ABB RAPID module: test.modx

MODULE A1_457_L
    ! ----------------------------------------------------------------------
    ! Robot ABB serial n. IRB  6720-101047
    ! ----------------------------------------------------------------------
    ! Final customer :  Martin Rea
    ! ----------------------------------------------------------------------
    ! Cell made by :    TREBI - Cellatica (BS) - Italy
    ! ----------------------------------------------------------------------
    ! Job order n. :    21301
    ! ----------------------------------------------------------------------
    ! Programmer :      Turati Simone
    ! ----------------------------------------------------------------------
    ! Date Rev.0:       07/10/2026
    ! Date Rev.1:
    ! Date Rev.2:
    ! Date Rev.3:
    ! Date Rev.4:
    ! ----------------------------------------------------------------------
    ! +-+-+-+-+-+-+-+-+-+-+-+-+-+-+-+-+-+-+-+-+-+-+-+-+-+-+-+-+-+-+-+-+-+-+-
    ! +-+-+-+-+-+-+-+-+-+-+-+-+-+-+-+-+-+-+-+-+-+-+-+-+-+-+-+-+-+-+-+-+-+-+-
    ! +-+-+-+-+-+-+-+-+-+-+-+-+-+-+-+-+-+-+-+-+-+-+-+-+-+-+-+-+-+-+-+-+-+-+-
    !EXCHANGE DATA (Variables with "M")
    ! **********************************************************************
    ! NUM DATA
    ! **********************************************************************
    PERS num nMProg:=1;
    ! **********************************************************************
    ! STRING DATA
    ! **********************************************************************
    !Stringhe nome programma
    PERS String sMProgramName:="PART_0001";
    PERS String sMPartName:="PEZZO 1";
    ! +-+-+-+-+-+-+-+-+-+-+-+-+-+-+-+-+-+-+-+-+-+-+-+-+-+-+-+-+-+-+-+-+-+-+-
    ! +-+-+-+-+-+-+-+-+-+-+-+-+-+-+-+-+-+-+-+-+-+-+-+-+-+-+-+-+-+-+-+-+-+-+-
    ! +-+-+-+-+-+-+-+-+-+-+-+-+-+-+-+-+-+-+-+-+-+-+-+-+-+-+-+-+-+-+-+-+-+-+-
    ! **********************************************************************
    ! NUM DATA
    ! **********************************************************************
    PERS dnum nLPartCounter:=19;
    ! **********************************************************************
    ! TOOL DATA
    ! **********************************************************************
    PERS tooldata tGripp_1:=[TRUE,[[0,250,335],[1,0,0,0]],[61.3,[54,3.3,163.7],[1,0,0,0],4.49,1.158,5.024]];
    ! **********************************************************************
    ! LOAD DATA
    ! **********************************************************************
    PERS loaddata LoadPart_L:=[4.5,[16.9,32.5,271],[1,0,0,0],0.7,0.6,0.2];
    ! **********************************************************************
    ! SPEED DATA
    ! **********************************************************************
    LOCAL PERS speeddata vPicking:=[60,500,0,0];
    LOCAL PERS speeddata vUnload:=[150,500,0,0];
    LOCAL PERS speeddata vGrind1:=[200,100,0,0];
    LOCAL PERS speeddata vGrind2:=[170,80,0,0];
    ! **********************************************************************
    ! ROBTARGET DATA
    ! **********************************************************************
    ! LOAD BELT
    PERS robtarget pLAppPick:=[[800,1370,1180],[0,0.642788,-0.766044,0],[0,0,-1,0],[9E+09,9E+09,9E+09,9E+09,9E+09,9E+09]];
    PERS robtarget pLPick:=[[3.81937,161.237,727.32],[0.138322,-0.983291,0.0782176,0.0888119],[0,-1,0,0],[9E+09,9E+09,9E+09,9E+09,9E+09,9E+09]];
    PERS robtarget pLPick_0:=[[97.94,1368.66,727.32],[0.160804,-0.644231,0.746958,-0.0340974],[0,-1,0,0],[9E+09,9E+09,9E+09,9E+09,9E+09,9E+09]];
    PERS robtarget pLCHK_Part:=[[-4.50,1321.99,1326.48],[0.156146,0.631329,-0.73609,-0.187653],[0,0,-1,0],[9E+09,9E+09,9E+09,9E+09,9E+09,9E+09]];
    ! RECENTRE
    PERS robtarget pLAppRec_:=[[890,-790,1800],[0,0,0.70711,-0.70711],[-1,-2,0,0],[9E+09,9E+09,9E+09,9E+09,9E+09,9E+09]];
    PERS robtarget pLRecentre_:=[[860,-495,2540],[0,0,0,1],[-1,-2,0,0],[9E+09,9E+09,9E+09,9E+09,9E+09,9E+09]];
    ! DATAMATRIX
    PERS robtarget pLAppDataMatrix_:=[[640.77,1371.32,1306.69],[0.400689,0.173653,-0.899217,0.0265008],[0,0,0,0],[9E+09,9E+09,9E+09,9E+09,9E+09,9E+09]];
    PERS robtarget pLDataMatrix:=[[-260,1005,1305],[0.407608,0.15668,-0.89732,0.0642135],[0,0,0,0],[9E+09,9E+09,9E+09,9E+09,9E+09,9E+09]];
    ! **********************************************************************
    ! CHANGE POINT
    PERS robtarget pLAppChange_1:=[[1370,1085,1560],[0,0,-0.707107,-0.707107],[0,1,-1,0],[9E+09,9E+09,9E+09,9E+09,9E+09,9E+09]];
    PERS robtarget pLAppChange_2:=[[1370,1085,1560],[0,0,-0.707107,-0.707107],[0,1,-1,0],[9E+09,9E+09,9E+09,9E+09,9E+09,9E+09]];
    PERS robtarget pLAppChange_3:=[[1370,1085,1560],[0,0,-0.707107,-0.707107],[0,1,-1,0],[9E+09,9E+09,9E+09,9E+09,9E+09,9E+09]];
    PERS robtarget pLAppChange_4:=[[1370,1085,1560],[0,0,-0.707107,-0.707107],[0,1,-1,0],[9E+09,9E+09,9E+09,9E+09,9E+09,9E+09]];
    PERS robtarget pLAppChange_5:=[[1370,1085,1560],[0,0,-0.707107,-0.707107],[0,1,-1,0],[9E+09,9E+09,9E+09,9E+09,9E+09,9E+09]];
    PERS robtarget pLAppChange_6:=[[1370,1085,1560],[0,0,-0.707107,-0.707107],[0,1,-1,0],[9E+09,9E+09,9E+09,9E+09,9E+09,9E+09]];
    PERS robtarget pLAppChange_7:=[[1370,1085,1560],[0,0,-0.707107,-0.707107],[0,1,-1,0],[9E+09,9E+09,9E+09,9E+09,9E+09,9E+09]];
    PERS robtarget pLAppChange_8:=[[1370,1085,1560],[0,0,-0.707107,-0.707107],[0,1,-1,0],[9E+09,9E+09,9E+09,9E+09,9E+09,9E+09]];
    PERS robtarget pLAppChange_9:=[[1370,1085,1560],[0,0,-0.707107,-0.707107],[0,1,-1,0],[9E+09,9E+09,9E+09,9E+09,9E+09,9E+09]];
    PERS robtarget pLAppChange_10:=[[1370,1085,1560],[0,0,-0.707107,-0.707107],[0,1,-1,0],[9E+09,9E+09,9E+09,9E+09,9E+09,9E+09]];
    PERS robtarget pLChange:=[[1590,1800,1695],[0,0,0.707107,0.707107],[0,1,-1,0],[9E+09,9E+09,9E+09,9E+09,9E+09,9E+09]];
    ! **********************************************************************
    !Safe Homing
    PERS robtarget pLSafeHoming_OP010_:=[[0,0,0],[0,0,0,0],[0,0,0,0],[9E+09,9E+09,9E+09,9E+09,9E+09,9E+09]];
    PERS robtarget pLSafeHoming_OP020_:=[[0,0,0],[0,0,0,0],[0,0,0,0],[9E+09,9E+09,9E+09,9E+09,9E+09,9E+09]];
    PERS robtarget pLSafeHoming_OP030_:=[[0,0,0],[0,0,0,0],[0,0,0,0],[9E+09,9E+09,9E+09,9E+09,9E+09,9E+09]];
    PERS robtarget pLSafeHoming_OP040_:=[[0,0,0],[0,0,0,0],[0,0,0,0],[9E+09,9E+09,9E+09,9E+09,9E+09,9E+09]];
    PERS robtarget pLSafeHoming_OP050_:=[[0,0,0],[0,0,0,0],[0,0,0,0],[9E+09,9E+09,9E+09,9E+09,9E+09,9E+09]];
    PERS robtarget pLSafeHoming_OP060_:=[[0,0,0],[0,0,0,0],[0,0,0,0],[9E+09,9E+09,9E+09,9E+09,9E+09,9E+09]];
    PERS robtarget pLSafeHoming_OP070_:=[[0,0,0],[0,0,0,0],[0,0,0,0],[9E+09,9E+09,9E+09,9E+09,9E+09,9E+09]];
    PERS robtarget pLSafeHoming_OP080_:=[[0,0,0],[0,0,0,0],[0,0,0,0],[9E+09,9E+09,9E+09,9E+09,9E+09,9E+09]];
    PERS robtarget pLSafeHoming_OP090_:=[[0,0,0],[0,0,0,0],[0,0,0,0],[9E+09,9E+09,9E+09,9E+09,9E+09,9E+09]];
    PERS robtarget pLSafeHoming_OP100_:=[[0,0,0],[0,0,0,0],[0,0,0,0],[9E+09,9E+09,9E+09,9E+09,9E+09,9E+09]];
    PERS robtarget pLSafeHoming_OP110_:=[[0,0,0],[0,0,0,0],[0,0,0,0],[9E+09,9E+09,9E+09,9E+09,9E+09,9E+09]];
    PERS robtarget pLSafeHoming_OP120_:=[[0,0,0],[0,0,0,0],[0,0,0,0],[9E+09,9E+09,9E+09,9E+09,9E+09,9E+09]];
    PERS robtarget pLSafeHoming_OP130_:=[[0,0,0],[0,0,0,0],[0,0,0,0],[9E+09,9E+09,9E+09,9E+09,9E+09,9E+09]];
    PERS robtarget pLSafeHoming_OP140_:=[[0,0,0],[0,0,0,0],[0,0,0,0],[9E+09,9E+09,9E+09,9E+09,9E+09,9E+09]];
    PERS robtarget pLSafeHoming_OP150_:=[[0,0,0],[0,0,0,0],[0,0,0,0],[9E+09,9E+09,9E+09,9E+09,9E+09,9E+09]];
    PERS robtarget pLSafeHoming_OP160_:=[[0,0,0],[0,0,0,0],[0,0,0,0],[9E+09,9E+09,9E+09,9E+09,9E+09,9E+09]];
    PERS robtarget pLSafeHoming_OP170_:=[[0,0,0],[0,0,0,0],[0,0,0,0],[9E+09,9E+09,9E+09,9E+09,9E+09,9E+09]];
    PERS robtarget pLSafeHoming_OP180_:=[[0,0,0],[0,0,0,0],[0,0,0,0],[9E+09,9E+09,9E+09,9E+09,9E+09,9E+09]];
    PERS robtarget pLSafeHoming_OP190_:=[[0,0,0],[0,0,0,0],[0,0,0,0],[9E+09,9E+09,9E+09,9E+09,9E+09,9E+09]];
    PERS robtarget pLSafeHoming_OP200_:=[[0,0,0],[0,0,0,0],[0,0,0,0],[9E+09,9E+09,9E+09,9E+09,9E+09,9E+09]];
    ! **********************************************************************
    ! GRINDER 1
    ! **********************************************************************
    !OPXXX
    PERS robtarget pLU1_OPXXX_000:=[[0,0,0],[0,0,0,0],[0,0,0,0],[9E+09,9E+09,9E+09,9E+09,9E+09,9E+09]];
    PERS robtarget pLU1_OPXXX_010:=[[0,0,0],[0,0,0,0],[0,0,0,0],[9E+09,9E+09,9E+09,9E+09,9E+09,9E+09]];
    PERS robtarget pLU1_OPXXX_020:=[[0,0,0],[0,0,0,0],[0,0,0,0],[9E+09,9E+09,9E+09,9E+09,9E+09,9E+09]];
    PERS robtarget pLU1_OPXXX_030:=[[0,0,0],[0,0,0,0],[0,0,0,0],[9E+09,9E+09,9E+09,9E+09,9E+09,9E+09]];
    ! **********************************************************************
    ! GRINDER 2
    ! **********************************************************************
    !OP10
    PERS robtarget pLU2_OP10_000 := [[-512.78,-45.67,-339.98],[0.753965,0.177077,0.558855,-0.296414],[-1,1,2,0],[9E+09,9E+09,9E+09,9E+09,9E+09,9E+09]];
    PERS robtarget pLU2_OP10_010 := [[83.19,99.41,-382.48],[0.834702,0.222849,0.429026,-0.263719],[-1,2,2,0],[9E+09,9E+09,9E+09,9E+09,9E+09,9E+09]];
    PERS robtarget pLU2_OP10_020 := [[166.56,99.41,-332.86],[0.834697,0.222853,0.429032,-0.26372],[-1,2,2,0],[9E+09,9E+09,9E+09,9E+09,9E+09,9E+09]];
    PERS robtarget pLU2_OP10_030 := [[166.56,99.41,-309.01],[0.834699,0.222852,0.42903,-0.26372],[-1,2,2,0],[9E+09,9E+09,9E+09,9E+09,9E+09,9E+09]];
    PERS robtarget pLU2_OP10_040 := [[147.76,53.29,-309.01],[0.834699,0.222851,0.429031,-0.26372],[-1,2,2,0],[9E+09,9E+09,9E+09,9E+09,9E+09,9E+09]];
    PERS robtarget pLU2_OP10_050 := [[99.74,9.11,-312.84],[0.834697,0.222851,0.429033,-0.26372],[-1,2,2,0],[9E+09,9E+09,9E+09,9E+09,9E+09,9E+09]];
    PERS robtarget pLU2_OP10_060 := [[89.03,-30.27,-311.48],[0.834674,0.222871,0.429035,-0.263775],[-1,2,2,0],[9E+09,9E+09,9E+09,9E+09,9E+09,9E+09]];
    PERS robtarget pLU2_OP10_070 := [[89.03,-66.46,-311.47],[0.834674,0.222871,0.429033,-0.263777],[-1,2,2,0],[9E+09,9E+09,9E+09,9E+09,9E+09,9E+09]];
    PERS robtarget pLU2_OP10_080 := [[78.00,-94.61,-311.47],[0.86058,0.168979,0.452974,-0.160198],[-1,1,2,0],[9E+09,9E+09,9E+09,9E+09,9E+09,9E+09]];
    PERS robtarget pLU2_OP10_090 := [[48.43,-125.73,-310.69],[0.86058,0.168979,0.452973,-0.160199],[-1,1,2,0],[9E+09,9E+09,9E+09,9E+09,9E+09,9E+09]];
    PERS robtarget pLU2_OP10_100 := [[48.68,-150.17,-329.57],[0.86058,0.168977,0.452973,-0.160199],[-1,1,2,0],[9E+09,9E+09,9E+09,9E+09,9E+09,9E+09]];
    PERS robtarget pLU2_OP10_110 := [[-99.73,-229.10,-399.55],[0.860581,0.168977,0.452973,-0.160199],[-1,1,2,0],[9E+09,9E+09,9E+09,9E+09,9E+09,9E+09]];
    !OP20
    PERS robtarget pLU2_OP20_000 := [[-385.23,300.06,-127.42],[0.574393,0.0777966,0.781268,-0.231604],[-1,1,2,0],[9E+09,9E+09,9E+09,9E+09,9E+09,9E+09]];
    PERS robtarget pLU2_OP20_010 := [[9.44,300.13,-103.22],[0.574395,0.0777988,0.781267,-0.231602],[-1,1,2,0],[9E+09,9E+09,9E+09,9E+09,9E+09,9E+09]];
    PERS robtarget pLU2_OP20_020 := [[101.46,300.12,-56.96],[0.574396,0.0778002,0.781266,-0.231603],[-1,1,2,0],[9E+09,9E+09,9E+09,9E+09,9E+09,9E+09]];
    PERS robtarget pLU2_OP20_030 := [[101.45,300.13,-43.36],[0.574393,0.0778009,0.781269,-0.231601],[-1,1,2,0],[9E+09,9E+09,9E+09,9E+09,9E+09,9E+09]];
    PERS robtarget pLU2_OP20_040 := [[101.45,261.09,-43.36],[0.574393,0.0778004,0.781269,-0.231601],[-1,1,2,0],[9E+09,9E+09,9E+09,9E+09,9E+09,9E+09]];
    PERS robtarget pLU2_OP20_050 := [[83.98,199.96,-132.65],[0.51864,-0.0749808,0.781563,-0.338452],[-1,1,1,0],[9E+09,9E+09,9E+09,9E+09,9E+09,9E+09]];
    PERS robtarget pLU2_OP20_060 := [[61.27,141.16,-169.72],[0.484154,-0.148838,0.770917,-0.386173],[-1,1,1,0],[9E+09,9E+09,9E+09,9E+09,9E+09,9E+09]];
    PERS robtarget pLU2_OP20_070 := [[8.24,67.49,-196.86],[0.423511,-0.258329,0.74142,-0.451886],[-1,1,1,0],[9E+09,9E+09,9E+09,9E+09,9E+09,9E+09]];
    PERS robtarget pLU2_OP20_080 := [[-7.60,-20.50,-212.03],[0.535292,-0.361141,0.639907,-0.416604],[-1,1,1,0],[9E+09,9E+09,9E+09,9E+09,9E+09,9E+09]];
    PERS robtarget pLU2_OP20_090 := [[30.73,-102.48,-219.34],[0.642287,-0.465548,0.487193,-0.365207],[-1,1,1,0],[9E+09,9E+09,9E+09,9E+09,9E+09,9E+09]];
    PERS robtarget pLU2_OP20_100 := [[-10.33,-244.75,-231.02],[0.642287,-0.465548,0.487193,-0.365206],[-1,1,1,0],[9E+09,9E+09,9E+09,9E+09,9E+09,9E+09]];
    PERS robtarget pLU2_OP20_110 := [[-10.33,-271.45,-231.03],[0.642288,-0.465548,0.487194,-0.365204],[-1,1,1,0],[9E+09,9E+09,9E+09,9E+09,9E+09,9E+09]];
    PERS robtarget pLU2_OP20_120 := [[-10.33,-292.72,-251.68],[0.642291,-0.465541,0.487206,-0.36519],[-1,1,1,0],[9E+09,9E+09,9E+09,9E+09,9E+09,9E+09]];
    PERS robtarget pLU2_OP20_130 := [[-190.07,-292.69,-351.19],[0.642289,-0.465559,0.48719,-0.365193],[-1,1,1,0],[9E+09,9E+09,9E+09,9E+09,9E+09,9E+09]];
    !OP30
    PERS robtarget pLU2_OP30_000 := [[-606.31,-417.45,-360.46],[0.0526328,0.614277,0.20406,0.76043],[-1,1,-1,0],[9E+09,9E+09,9E+09,9E+09,9E+09,9E+09]];
    PERS robtarget pLU2_OP30_010 := [[-17.06,-336.23,-338.16],[0.0526321,0.614273,0.204057,0.760433],[-1,1,0,0],[9E+09,9E+09,9E+09,9E+09,9E+09,9E+09]];
    PERS robtarget pLU2_OP30_020 := [[52.21,-336.22,-282.57],[0.0526289,0.614275,0.204054,0.760433],[-1,1,0,0],[9E+09,9E+09,9E+09,9E+09,9E+09,9E+09]];
    PERS robtarget pLU2_OP30_030 := [[52.06,-318.83,-265.48],[0.0526342,0.614272,0.204059,0.760434],[-1,1,0,0],[9E+09,9E+09,9E+09,9E+09,9E+09,9E+09]];
    PERS robtarget pLU2_OP30_040 := [[52.06,-288.05,-265.48],[0.0526341,0.614272,0.204059,0.760434],[-1,1,0,0],[9E+09,9E+09,9E+09,9E+09,9E+09,9E+09]];
    PERS robtarget pLU2_OP30_050 := [[52.06,-258.93,-255.88],[0.052635,0.614272,0.204059,0.760434],[-1,1,0,0],[9E+09,9E+09,9E+09,9E+09,9E+09,9E+09]];
    PERS robtarget pLU2_OP30_060 := [[60.46,-173.47,-251.63],[0.0526278,0.614276,0.204056,0.760431],[-1,1,0,0],[9E+09,9E+09,9E+09,9E+09,9E+09,9E+09]];
    PERS robtarget pLU2_OP30_070 := [[60.46,-162.14,-250.24],[0.0526281,0.614276,0.204057,0.760432],[-1,1,0,0],[9E+09,9E+09,9E+09,9E+09,9E+09,9E+09]];
    PERS robtarget pLU2_OP30_080 := [[72.17,-150.18,-228.58],[0.0526243,0.614279,0.204054,0.76043],[-1,1,0,0],[9E+09,9E+09,9E+09,9E+09,9E+09,9E+09]];
    PERS robtarget pLU2_OP30_090 := [[72.19,-115.25,-231.76],[0.0526317,0.614273,0.204059,0.760433],[-1,1,0,0],[9E+09,9E+09,9E+09,9E+09,9E+09,9E+09]];
    PERS robtarget pLU2_OP30_100 := [[73.88,-65.85,-234.90],[0.0526266,0.614276,0.204058,0.760432],[-1,1,0,0],[9E+09,9E+09,9E+09,9E+09,9E+09,9E+09]];
    PERS robtarget pLU2_OP30_110 := [[73.93,-33.88,-234.89],[0.0526271,0.614275,0.204058,0.760432],[-1,1,0,0],[9E+09,9E+09,9E+09,9E+09,9E+09,9E+09]];
    PERS robtarget pLU2_OP30_120 := [[88.72,-11.35,-221.02],[0.0526255,0.614275,0.20406,0.760432],[-1,1,0,0],[9E+09,9E+09,9E+09,9E+09,9E+09,9E+09]];
    PERS robtarget pLU2_OP30_130 := [[100.68,56.41,-214.86],[0.00740228,-0.617052,-0.128267,-0.776363],[-1,1,0,0],[9E+09,9E+09,9E+09,9E+09,9E+09,9E+09]];
    PERS robtarget pLU2_OP30_140 := [[100.68,135.16,-185.77],[0.0962711,-0.609235,-0.0190289,-0.786894],[-1,1,0,0],[9E+09,9E+09,9E+09,9E+09,9E+09,9E+09]];
    PERS robtarget pLU2_OP30_150 := [[100.66,173.20,-160.73],[0.14348,-0.601643,0.0462119,-0.784413],[-1,1,0,0],[9E+09,9E+09,9E+09,9E+09,9E+09,9E+09]];
    PERS robtarget pLU2_OP30_160 := [[100.69,199.74,-135.33],[0.178665,-0.590179,0.105027,-0.780216],[-1,1,0,0],[9E+09,9E+09,9E+09,9E+09,9E+09,9E+09]];
    PERS robtarget pLU2_OP30_170 := [[101.34,338.20,-122.10],[0.178664,-0.590171,0.10502,-0.780223],[-1,1,0,0],[9E+09,9E+09,9E+09,9E+09,9E+09,9E+09]];
    PERS robtarget pLU2_OP30_180 := [[101.82,359.38,-120.37],[0.178667,-0.590179,0.105026,-0.780216],[-1,1,0,0],[9E+09,9E+09,9E+09,9E+09,9E+09,9E+09]];
    PERS robtarget pLU2_OP30_190 := [[101.82,370.03,-117.04],[0.178666,-0.590176,0.105022,-0.780218],[-1,1,0,0],[9E+09,9E+09,9E+09,9E+09,9E+09,9E+09]];
    PERS robtarget pLU2_OP30_200 := [[102.02,378.40,-82.10],[0.178665,-0.590174,0.105021,-0.78022],[-1,1,0,0],[9E+09,9E+09,9E+09,9E+09,9E+09,9E+09]];
    PERS robtarget pLU2_OP30_210 := [[102.03,422.66,-82.10],[0.178665,-0.590173,0.105021,-0.780221],[-1,1,0,0],[9E+09,9E+09,9E+09,9E+09,9E+09,9E+09]];
    PERS robtarget pLU2_OP30_220 := [[102.44,480.96,-82.10],[0.178665,-0.590174,0.105022,-0.78022],[0,1,0,0],[9E+09,9E+09,9E+09,9E+09,9E+09,9E+09]];
    PERS robtarget pLU2_OP30_230 := [[102.43,480.20,96.79],[0.178665,-0.59017,0.105018,-0.780224],[0,1,0,0],[9E+09,9E+09,9E+09,9E+09,9E+09,9E+09]];
    PERS robtarget pLU2_OP30_240 := [[161.68,397.29,2.47],[0.0655787,-0.702265,0.137697,-0.695386],[0,1,0,0],[9E+09,9E+09,9E+09,9E+09,9E+09,9E+09]];
    PERS robtarget pLU2_OP30_250 := [[161.69,397.29,2.49],[0.0655788,-0.702262,0.137697,-0.69539],[0,1,0,0],[9E+09,9E+09,9E+09,9E+09,9E+09,9E+09]];
    PERS robtarget pLU2_OP30_260 := [[161.69,415.52,2.48],[0.065579,-0.702264,0.137698,-0.695388],[0,1,0,0],[9E+09,9E+09,9E+09,9E+09,9E+09,9E+09]];
    PERS robtarget pLU2_OP30_270 := [[161.69,428.24,21.00],[0.0655789,-0.702263,0.137697,-0.695389],[0,1,0,0],[9E+09,9E+09,9E+09,9E+09,9E+09,9E+09]];
    PERS robtarget pLU2_OP30_280 := [[162.84,611.07,21.00],[0.0655725,-0.702264,0.137706,-0.695387],[0,2,0,0],[9E+09,9E+09,9E+09,9E+09,9E+09,9E+09]];
    PERS robtarget pLU2_OP30_290 := [[96.32,76.93,-471.17],[0.559851,0.638465,0.232535,0.474191],[-1,2,-1,0],[9E+09,9E+09,9E+09,9E+09,9E+09,9E+09]];
    PERS robtarget pLU2_OP30_300 := [[95.34,-11.04,-420.70],[0.559851,0.638464,0.232536,0.474191],[-1,1,-1,0],[9E+09,9E+09,9E+09,9E+09,9E+09,9E+09]];
    PERS robtarget pLU2_OP30_310 := [[95.33,-16.30,-406.32],[0.559852,0.638464,0.232534,0.474191],[-1,1,-1,0],[9E+09,9E+09,9E+09,9E+09,9E+09,9E+09]];
    PERS robtarget pLU2_OP30_320 := [[95.33,8.06,-406.32],[0.559852,0.638464,0.232535,0.474191],[-1,1,-1,0],[9E+09,9E+09,9E+09,9E+09,9E+09,9E+09]];
    PERS robtarget pLU2_OP30_330 := [[95.31,8.03,-422.81],[0.559852,0.63847,0.232533,0.474183],[-1,1,-1,0],[9E+09,9E+09,9E+09,9E+09,9E+09,9E+09]];
    PERS robtarget pLU2_OP30_340 := [[113.89,8.35,-458.89],[0.482927,0.600997,0.321749,0.549602],[-1,1,-1,0],[9E+09,9E+09,9E+09,9E+09,9E+09,9E+09]];
    PERS robtarget pLU2_OP30_350 := [[113.89,-33.86,-435.57],[0.482928,0.600995,0.321751,0.549602],[-1,1,-1,0],[9E+09,9E+09,9E+09,9E+09,9E+09,9E+09]];
    PERS robtarget pLU2_OP30_360 := [[104.34,-56.68,-435.57],[0.482926,0.600995,0.321751,0.549603],[-1,1,-1,0],[9E+09,9E+09,9E+09,9E+09,9E+09,9E+09]];
    PERS robtarget pLU2_OP30_370 := [[97.09,-80.58,-439.37],[0.429334,0.578514,0.370309,0.586401],[-1,1,-1,0],[9E+09,9E+09,9E+09,9E+09,9E+09,9E+09]];
    PERS robtarget pLU2_OP30_380 := [[84.59,-111.35,-432.91],[0.429335,0.578511,0.37031,0.586402],[-1,1,-1,0],[9E+09,9E+09,9E+09,9E+09,9E+09,9E+09]];
    PERS robtarget pLU2_OP30_390 := [[84.59,-132.56,-440.51],[0.429339,0.578508,0.370309,0.586402],[-1,1,-1,0],[9E+09,9E+09,9E+09,9E+09,9E+09,9E+09]];
    PERS robtarget pLU2_OP30_400 := [[84.60,-134.22,-394.80],[0.429346,0.578494,0.370319,0.586405],[-1,1,-1,0],[9E+09,9E+09,9E+09,9E+09,9E+09,9E+09]];
    PERS robtarget pLU2_OP30_410 := [[84.60,-124.72,-373.35],[0.429346,0.578494,0.370317,0.586406],[-1,1,-1,0],[9E+09,9E+09,9E+09,9E+09,9E+09,9E+09]];
    PERS robtarget pLU2_OP30_420 := [[84.60,-146.35,-373.35],[0.429345,0.578494,0.370318,0.586406],[-1,1,-1,0],[9E+09,9E+09,9E+09,9E+09,9E+09,9E+09]];
    PERS robtarget pLU2_OP30_430 := [[84.61,-173.54,-373.34],[0.429351,0.578489,0.370317,0.586407],[-1,1,-1,0],[9E+09,9E+09,9E+09,9E+09,9E+09,9E+09]];
    PERS robtarget pLU2_OP30_440 := [[-10.13,-222.88,-433.94],[0.429346,0.578494,0.370317,0.586406],[-1,1,-1,0],[9E+09,9E+09,9E+09,9E+09,9E+09,9E+09]];
    !OP70
    PERS robtarget pLU2_OP070_000:=[[-408.28,-45.28,414.95],[0.437495,-0.259727,0.675398,-0.533833],[-1,0,2,0],[9E+09,9E+09,9E+09,9E+09,9E+09,9E+09]];
    PERS robtarget pLU2_OP070_010:=[[-72.80,61.79,414.96],[0.437497,-0.259728,0.675394,-0.533837],[-1,0,2,0],[9E+09,9E+09,9E+09,9E+09,9E+09,9E+09]];
    PERS robtarget pLU2_OP070_020:=[[64.33,61.81,414.89],[0.437487,-0.25973,0.675405,-0.533828],[-1,0,2,0],[9E+09,9E+09,9E+09,9E+09,9E+09,9E+09]];
    PERS robtarget pLU2_OP070_030:=[[70.54,61.79,400.67],[0.437496,-0.259729,0.675392,-0.533838],[-1,1,2,0],[9E+09,9E+09,9E+09,9E+09,9E+09,9E+09]];
    PERS robtarget pLU2_OP070_040:=[[72.42,66.18,357.75],[0.437497,-0.259728,0.67539,-0.533841],[-1,1,1,0],[9E+09,9E+09,9E+09,9E+09,9E+09,9E+09]];
    PERS robtarget pLU2_OP070_050:=[[73.32,77.42,345.41],[0.437497,-0.259727,0.675391,-0.53384],[-1,1,1,0],[9E+09,9E+09,9E+09,9E+09,9E+09,9E+09]];
    PERS robtarget pLU2_OP070_060:=[[72.97,77.43,337.09],[0.440655,-0.263725,0.673837,-0.531239],[-1,1,1,0],[9E+09,9E+09,9E+09,9E+09,9E+09,9E+09]];
    PERS robtarget pLU2_OP070_070:=[[73.94,79.71,316.54],[0.440658,-0.263725,0.673834,-0.531242],[-1,1,1,0],[9E+09,9E+09,9E+09,9E+09,9E+09,9E+09]];
    PERS robtarget pLU2_OP070_080:=[[69.94,83.17,310.35],[0.440657,-0.263725,0.673835,-0.531241],[-1,1,1,0],[9E+09,9E+09,9E+09,9E+09,9E+09,9E+09]];
    PERS robtarget pLU2_OP070_090:=[[-528.55,83.17,310.34],[0.440657,-0.263724,0.673837,-0.531239],[-1,0,2,0],[9E+09,9E+09,9E+09,9E+09,9E+09,9E+09]];
    !OP80
    PERS robtarget pLU2_OP080_000:=[[-439.18,139.36,266.67],[0.237607,-0.308213,0.546191,-0.741771],[-1,2,0,0],[9E+09,9E+09,9E+09,9E+09,9E+09,9E+09]];
    PERS robtarget pLU2_OP080_010:=[[-14.57,129.75,2.02],[0.237605,-0.308215,0.546193,-0.741769],[-1,2,0,0],[9E+09,9E+09,9E+09,9E+09,9E+09,9E+09]];
    PERS robtarget pLU2_OP080_020:=[[93.51,129.75,-16.65],[0.237606,-0.30821,0.546192,-0.741771],[-1,2,0,0],[9E+09,9E+09,9E+09,9E+09,9E+09,9E+09]];
    PERS robtarget pLU2_OP080_030:=[[104.86,129.75,-29.48],[0.237608,-0.308212,0.546191,-0.74177],[-1,2,0,0],[9E+09,9E+09,9E+09,9E+09,9E+09,9E+09]];
    PERS robtarget pLU2_OP080_040:=[[102.67,129.75,-61.93],[0.237608,-0.308214,0.54619,-0.74177],[-1,2,0,0],[9E+09,9E+09,9E+09,9E+09,9E+09,9E+09]];
    PERS robtarget pLU2_OP080_050:=[[97.60,129.75,-69.46],[0.237608,-0.30821,0.54619,-0.741772],[-1,2,0,0],[9E+09,9E+09,9E+09,9E+09,9E+09,9E+09]];
    PERS robtarget pLU2_OP080_060:=[[-392.81,209.79,-69.46],[0.237608,-0.308211,0.546189,-0.741772],[-1,2,0,0],[9E+09,9E+09,9E+09,9E+09,9E+09,9E+09]];
    !OP90
    PERS robtarget pLU2_OP090_000:=[[-496.10,203.40,-54.83],[0.251573,-0.284697,0.494783,-0.781568],[-1,2,0,0],[9E+09,9E+09,9E+09,9E+09,9E+09,9E+09]];
    PERS robtarget pLU2_OP090_010:=[[1.29,190.38,-154.04],[0.251575,-0.284694,0.49478,-0.78157],[0,2,0,0],[9E+09,9E+09,9E+09,9E+09,9E+09,9E+09]];
    PERS robtarget pLU2_OP090_020:=[[111.05,140.40,-154.06],[0.251572,-0.284698,0.494785,-0.781567],[-1,2,0,0],[9E+09,9E+09,9E+09,9E+09,9E+09,9E+09]];
    PERS robtarget pLU2_OP090_030:=[[120.67,140.40,-171.46],[0.251569,-0.284702,0.494787,-0.781565],[-1,2,0,0],[9E+09,9E+09,9E+09,9E+09,9E+09,9E+09]];
    PERS robtarget pLU2_OP090_040:=[[118.92,140.38,-201.03],[0.251563,-0.284695,0.494792,-0.781566],[-1,2,0,0],[9E+09,9E+09,9E+09,9E+09,9E+09,9E+09]];
    PERS robtarget pLU2_OP090_050:=[[114.86,140.37,-215.26],[0.251563,-0.284695,0.494793,-0.781565],[-1,2,0,0],[9E+09,9E+09,9E+09,9E+09,9E+09,9E+09]];
    PERS robtarget pLU2_OP090_060:=[[-409.57,230.34,-215.25],[0.251565,-0.284694,0.49479,-0.781567],[-1,2,0,0],[9E+09,9E+09,9E+09,9E+09,9E+09,9E+09]];
    !OP100
    PERS robtarget pLU2_OP100_000:=[[-470.91,154.77,-154.01],[0.314743,-0.352653,0.421479,-0.773905],[-1,1,0,0],[9E+09,9E+09,9E+09,9E+09,9E+09,9E+09]];
    PERS robtarget pLU2_OP100_010:=[[-3.88,154.76,-259.09],[0.314737,-0.35266,0.421493,-0.773896],[-1,2,0,0],[9E+09,9E+09,9E+09,9E+09,9E+09,9E+09]];
    PERS robtarget pLU2_OP100_020:=[[102.60,154.76,-256.29],[0.314739,-0.35266,0.421492,-0.773896],[-1,2,0,0],[9E+09,9E+09,9E+09,9E+09,9E+09,9E+09]];
    PERS robtarget pLU2_OP100_030:=[[110.15,154.76,-253.29],[0.31474,-0.352656,0.421489,-0.773898],[-1,2,0,0],[9E+09,9E+09,9E+09,9E+09,9E+09,9E+09]];
    PERS robtarget pLU2_OP100_040:=[[110.16,154.74,-266.91],[0.314737,-0.352658,0.421497,-0.773895],[-1,2,0,0],[9E+09,9E+09,9E+09,9E+09,9E+09,9E+09]];
    PERS robtarget pLU2_OP100_050:=[[90.81,154.74,-266.90],[0.314738,-0.352656,0.421495,-0.773896],[-1,2,0,0],[9E+09,9E+09,9E+09,9E+09,9E+09,9E+09]];
    PERS robtarget pLU2_OP100_060:=[[-328.17,168.91,-266.92],[0.314737,-0.352659,0.421498,-0.773894],[-1,1,0,0],[9E+09,9E+09,9E+09,9E+09,9E+09,9E+09]];
    !OP110
    PERS robtarget pLU2_OP110_000:=[[-349.31,177.69,-267.83],[0.31474,-0.352642,0.421491,-0.773904],[-1,1,0,0],[9E+09,9E+09,9E+09,9E+09,9E+09,9E+09]];
    PERS robtarget pLU2_OP110_010:=[[13.19,177.70,-267.83],[0.314741,-0.352641,0.421489,-0.773905],[-1,2,0,0],[9E+09,9E+09,9E+09,9E+09,9E+09,9E+09]];
    PERS robtarget pLU2_OP110_020:=[[99.49,177.69,-267.79],[0.314745,-0.352635,0.421479,-0.773912],[-1,2,0,0],[9E+09,9E+09,9E+09,9E+09,9E+09,9E+09]];
    PERS robtarget pLU2_OP110_030:=[[110.86,177.69,-267.83],[0.31474,-0.352642,0.421489,-0.773905],[-1,2,0,0],[9E+09,9E+09,9E+09,9E+09,9E+09,9E+09]];
    PERS robtarget pLU2_OP110_040:=[[112.27,177.66,-304.50],[0.314734,-0.35264,0.421495,-0.773906],[-1,2,0,0],[9E+09,9E+09,9E+09,9E+09,9E+09,9E+09]];
    PERS robtarget pLU2_OP110_050:=[[101.82,177.66,-314.04],[0.314734,-0.352639,0.421494,-0.773906],[-1,2,0,0],[9E+09,9E+09,9E+09,9E+09,9E+09,9E+09]];
    PERS robtarget pLU2_OP110_060:=[[106.98,160.22,-272.46],[0.314725,-0.352637,0.421505,-0.773905],[-1,2,0,0],[9E+09,9E+09,9E+09,9E+09,9E+09,9E+09]];
    PERS robtarget pLU2_OP110_070:=[[111.57,160.19,-272.44],[0.314722,-0.352631,0.421505,-0.773909],[-1,2,0,0],[9E+09,9E+09,9E+09,9E+09,9E+09,9E+09]];
    PERS robtarget pLU2_OP110_080:=[[111.76,157.10,-289.24],[0.314726,-0.352638,0.421503,-0.773905],[-1,2,0,0],[9E+09,9E+09,9E+09,9E+09,9E+09,9E+09]];
    PERS robtarget pLU2_OP110_090:=[[115.09,144.85,-294.53],[0.308469,-0.349223,0.424334,-0.776422],[-1,2,0,0],[9E+09,9E+09,9E+09,9E+09,9E+09,9E+09]];
    PERS robtarget pLU2_OP110_100:=[[115.66,140.13,-305.05],[0.30847,-0.349223,0.424334,-0.776422],[-1,2,0,0],[9E+09,9E+09,9E+09,9E+09,9E+09,9E+09]];
    PERS robtarget pLU2_OP110_110:=[[110.78,140.13,-312.62],[0.308467,-0.349226,0.424336,-0.77642],[-1,2,0,0],[9E+09,9E+09,9E+09,9E+09,9E+09,9E+09]];
    PERS robtarget pLU2_OP110_120:=[[-381.10,140.13,-265.15],[0.30847,-0.349228,0.424338,-0.776417],[-1,1,0,0],[9E+09,9E+09,9E+09,9E+09,9E+09,9E+09]];
    !OP120
    PERS robtarget pLU2_OP120_000:=[[-454.64,-330.43,2.81],[0.084778,-0.685941,-0.24412,-0.680223],[-1,0,0,0],[9E+09,9E+09,9E+09,9E+09,9E+09,9E+09]];
    PERS robtarget pLU2_OP120_010:=[[-91.29,-330.42,2.81],[0.0847798,-0.685941,-0.244118,-0.680223],[-1,0,0,0],[9E+09,9E+09,9E+09,9E+09,9E+09,9E+09]];
    PERS robtarget pLU2_OP120_020:=[[35.15,-330.43,2.80],[0.0847826,-0.685942,-0.244116,-0.680223],[-1,1,0,0],[9E+09,9E+09,9E+09,9E+09,9E+09,9E+09]];
    PERS robtarget pLU2_OP120_030:=[[40.86,-330.43,2.80],[0.0847822,-0.685943,-0.244116,-0.680222],[-1,1,0,0],[9E+09,9E+09,9E+09,9E+09,9E+09,9E+09]];
    PERS robtarget pLU2_OP120_040:=[[77.18,-337.42,-49.36],[0.084781,-0.685941,-0.244119,-0.680222],[-1,1,0,0],[9E+09,9E+09,9E+09,9E+09,9E+09,9E+09]];
    PERS robtarget pLU2_OP120_050:=[[77.18,-337.42,-57.08],[0.0847805,-0.685941,-0.24412,-0.680222],[-1,1,0,0],[9E+09,9E+09,9E+09,9E+09,9E+09,9E+09]];
    PERS robtarget pLU2_OP120_060:=[[-499.44,-337.42,-57.09],[0.0847849,-0.685944,-0.244115,-0.680221],[-1,0,0,0],[9E+09,9E+09,9E+09,9E+09,9E+09,9E+09]];
    !OP130
    PERS robtarget pLU2_OP130_000:=[[-471.27,-260.06,12.19],[0.00880666,-0.601736,-0.293995,-0.742565],[-1,0,0,0],[9E+09,9E+09,9E+09,9E+09,9E+09,9E+09]];
    PERS robtarget pLU2_OP130_010:=[[-22.82,-260.04,12.19],[0.00881128,-0.601736,-0.293996,-0.742564],[-1,1,0,0],[9E+09,9E+09,9E+09,9E+09,9E+09,9E+09]];
    PERS robtarget pLU2_OP130_020:=[[44.25,-260.07,12.18],[0.00881067,-0.601738,-0.293994,-0.742564],[-1,1,0,0],[9E+09,9E+09,9E+09,9E+09,9E+09,9E+09]];
    PERS robtarget pLU2_OP130_030:=[[57.64,-260.05,12.21],[0.00881165,-0.601731,-0.293998,-0.742568],[-1,1,0,0],[9E+09,9E+09,9E+09,9E+09,9E+09,9E+09]];
    PERS robtarget pLU2_OP130_040:=[[45.01,-265.93,-13.85],[0.00880896,-0.601736,-0.293997,-0.742565],[-1,1,0,0],[9E+09,9E+09,9E+09,9E+09,9E+09,9E+09]];
    PERS robtarget pLU2_OP130_050:=[[37.08,-273.31,-29.22],[0.00882285,-0.601738,-0.294003,-0.74256],[-1,1,0,0],[9E+09,9E+09,9E+09,9E+09,9E+09,9E+09]];
    PERS robtarget pLU2_OP130_060:=[[18.45,-273.31,-70.36],[0.0088239,-0.60174,-0.294006,-0.742557],[-1,1,0,0],[9E+09,9E+09,9E+09,9E+09,9E+09,9E+09]];
    PERS robtarget pLU2_OP130_070:=[[2.14,-273.30,-70.36],[0.00882502,-0.60174,-0.294006,-0.742557],[-1,1,0,0],[9E+09,9E+09,9E+09,9E+09,9E+09,9E+09]];
    PERS robtarget pLU2_OP130_080:=[[-475.18,-270.85,-70.37],[0.00882762,-0.60174,-0.294006,-0.742557],[-1,0,0,0],[9E+09,9E+09,9E+09,9E+09,9E+09,9E+09]];
    !OP140
    PERS robtarget pLU2_OP140_000:=[[-594.58,-55.34,99.52],[0.00427089,0.828798,-0.20634,0.520096],[-1,0,1,0],[9E+09,9E+09,9E+09,9E+09,9E+09,9E+09]];
    PERS robtarget pLU2_OP140_010:=[[-180.62,-62.86,99.55],[0.00427237,0.828795,-0.206338,0.5201],[-1,0,1,0],[9E+09,9E+09,9E+09,9E+09,9E+09,9E+09]];
    PERS robtarget pLU2_OP140_020:=[[-54.97,-62.87,82.37],[0.0042716,0.828798,-0.206341,0.520096],[-1,0,1,0],[9E+09,9E+09,9E+09,9E+09,9E+09,9E+09]];
    PERS robtarget pLU2_OP140_030:=[[-45.84,-70.51,71.22],[0.00426719,0.828801,-0.206344,0.520089],[-1,0,1,0],[9E+09,9E+09,9E+09,9E+09,9E+09,9E+09]];
    PERS robtarget pLU2_OP140_040:=[[-41.96,-68.84,40.46],[0.00426893,0.8288,-0.206343,0.520092],[-1,0,1,0],[9E+09,9E+09,9E+09,9E+09,9E+09,9E+09]];
    PERS robtarget pLU2_OP140_050:=[[-41.60,-60.78,38.77],[0.0042701,0.828797,-0.206341,0.520097],[-1,0,1,0],[9E+09,9E+09,9E+09,9E+09,9E+09,9E+09]];
    PERS robtarget pLU2_OP140_060:=[[-38.69,-47.38,25.23],[0.00426723,0.828802,-0.206341,0.520089],[-1,0,1,0],[9E+09,9E+09,9E+09,9E+09,9E+09,9E+09]];
    PERS robtarget pLU2_OP140_070:=[[-48.73,-47.40,21.55],[0.00426969,0.828798,-0.206342,0.520094],[-1,0,1,0],[9E+09,9E+09,9E+09,9E+09,9E+09,9E+09]];
    PERS robtarget pLU2_OP140_080:=[[-553.87,-47.38,21.58],[0.0042773,0.828795,-0.206337,0.520101],[-1,0,1,0],[9E+09,9E+09,9E+09,9E+09,9E+09,9E+09]];
    !OP150
    PERS robtarget pLU2_OP150_000:=[[-552.85,97.78,-79.41],[0.381551,-0.215901,0.496414,-0.749252],[-1,1,1,0],[9E+09,9E+09,9E+09,9E+09,9E+09,9E+09]];
    PERS robtarget pLU2_OP150_010:=[[-38.02,93.70,-79.40],[0.381552,-0.215899,0.496413,-0.749253],[-1,2,0,0],[9E+09,9E+09,9E+09,9E+09,9E+09,9E+09]];
    PERS robtarget pLU2_OP150_020:=[[50.75,93.56,-79.39],[0.381553,-0.215895,0.496411,-0.749254],[-1,2,0,0],[9E+09,9E+09,9E+09,9E+09,9E+09,9E+09]];
    PERS robtarget pLU2_OP150_030:=[[56.55,93.56,-87.02],[0.381551,-0.2159,0.496416,-0.749251],[-1,2,0,0],[9E+09,9E+09,9E+09,9E+09,9E+09,9E+09]];
    PERS robtarget pLU2_OP150_040:=[[54.63,83.92,-124.10],[0.38154,-0.215901,0.49643,-0.749247],[-1,2,0,0],[9E+09,9E+09,9E+09,9E+09,9E+09,9E+09]];
    PERS robtarget pLU2_OP150_050:=[[47.41,83.92,-133.18],[0.38154,-0.215901,0.496429,-0.749248],[-1,2,0,0],[9E+09,9E+09,9E+09,9E+09,9E+09,9E+09]];
    PERS robtarget pLU2_OP150_060:=[[-460.80,83.92,-133.19],[0.381538,-0.215902,0.496433,-0.749246],[-1,1,1,0],[9E+09,9E+09,9E+09,9E+09,9E+09,9E+09]];
    !OP390
    PERS robtarget pLU2_OP390_000 := [[-550.18,111.81,-26.27],[0.313663,-0.103311,0.754315,-0.567407],[-1,2,0,0],[9E+09,9E+09,9E+09,9E+09,9E+09,9E+09]];
    PERS robtarget pLU2_OP390_010 := [[-30.08,111.80,-26.25],[0.313665,-0.10331,0.754312,-0.56741],[-1,2,0,0],[9E+09,9E+09,9E+09,9E+09,9E+09,9E+09]];
    PERS robtarget pLU2_OP390_020 := [[39.74,81.28,-26.21],[0.313673,-0.103304,0.754306,-0.567415],[-1,2,0,0],[9E+09,9E+09,9E+09,9E+09,9E+09,9E+09]];
    PERS robtarget pLU2_OP390_030 := [[45.80,81.27,-45.75],[0.313666,-0.10331,0.754311,-0.567412],[-1,2,0,0],[9E+09,9E+09,9E+09,9E+09,9E+09,9E+09]];
    PERS robtarget pLU2_OP390_040 := [[46.69,86.94,-79.36],[0.311906,-0.10199,0.755039,-0.567651],[-1,2,0,0],[9E+09,9E+09,9E+09,9E+09,9E+09,9E+09]];
    PERS robtarget pLU2_OP390_050 := [[44.15,97.02,-86.04],[0.311906,-0.10199,0.75504,-0.567651],[-1,2,0,0],[9E+09,9E+09,9E+09,9E+09,9E+09,9E+09]];
    PERS robtarget pLU2_OP390_060 := [[7.61,116.43,-86.05],[0.311904,-0.101992,0.75504,-0.567651],[-1,2,0,0],[9E+09,9E+09,9E+09,9E+09,9E+09,9E+09]];
    PERS robtarget pLU2_OP390_070 := [[38.51,-124.67,-191.60],[0.197261,-0.467763,0.0495327,-0.860135],[-1,1,0,0],[9E+09,9E+09,9E+09,9E+09,9E+09,9E+09]];
    PERS robtarget pLU2_OP390_080 := [[38.51,-124.67,-191.59],[0.197263,-0.467762,0.0495308,-0.860135],[-1,1,0,0],[9E+09,9E+09,9E+09,9E+09,9E+09,9E+09]];
    PERS robtarget pLU2_OP390_090 := [[16.42,173.24,-135.95],[0.465073,-0.277041,0.583178,-0.605688],[-1,1,1,0],[9E+09,9E+09,9E+09,9E+09,9E+09,9E+09]];
    PERS robtarget pLU2_OP390_100 := [[-830.91,-35.64,-68.30],[0.640247,-0.475858,0.562925,-0.216237],[-1,0,2,0],[9E+09,9E+09,9E+09,9E+09,9E+09,9E+09]];
    PERS robtarget pLU2_OP390_110 := [[-214.77,48.14,-68.32],[0.73606,-0.5117,0.427574,-0.116445],[-1,1,2,0],[9E+09,9E+09,9E+09,9E+09,9E+09,9E+09]];
    PERS robtarget pLU2_OP390_120 := [[-191.44,72.95,-68.31],[0.73606,-0.511702,0.427571,-0.116447],[-1,1,2,0],[9E+09,9E+09,9E+09,9E+09,9E+09,9E+09]];
    PERS robtarget pLU2_OP390_130 := [[-187.21,81.95,-80.40],[0.736064,-0.511697,0.42757,-0.116448],[-1,1,1,0],[9E+09,9E+09,9E+09,9E+09,9E+09,9E+09]];
    PERS robtarget pLU2_OP390_140 := [[-186.81,81.95,-98.10],[0.736064,-0.511698,0.427568,-0.116448],[-1,1,1,0],[9E+09,9E+09,9E+09,9E+09,9E+09,9E+09]];
    PERS robtarget pLU2_OP390_150 := [[-197.86,81.95,-110.44],[0.736065,-0.511693,0.427574,-0.116441],[-1,1,1,0],[9E+09,9E+09,9E+09,9E+09,9E+09,9E+09]];
    PERS robtarget pLU2_OP390_160 := [[-301.52,63.17,-110.42],[0.736064,-0.511697,0.427569,-0.116448],[-1,0,1,0],[9E+09,9E+09,9E+09,9E+09,9E+09,9E+09]];
    PERS robtarget pLU2_OP390_170 := [[-624.49,-66.79,-110.42],[0.736064,-0.511698,0.427569,-0.116449],[-1,0,1,0],[9E+09,9E+09,9E+09,9E+09,9E+09,9E+09]];
    !OP410
    PERS robtarget pLU2_OP410_000 := [[-594.58,-55.34,99.51],[0.00426986,0.828798,-0.206341,0.520094],[-1,0,1,0],[9E+09,9E+09,9E+09,9E+09,9E+09,9E+09]];
    PERS robtarget pLU2_OP410_010 := [[-219.14,-85.05,185.35],[0.12854,-0.701384,0.295207,-0.635917],[-1,1,1,0],[9E+09,9E+09,9E+09,9E+09,9E+09,9E+09]];
    PERS robtarget pLU2_OP410_020 := [[-138.62,-85.04,185.32],[0.128545,-0.701388,0.295211,-0.635911],[-1,1,1,0],[9E+09,9E+09,9E+09,9E+09,9E+09,9E+09]];
    PERS robtarget pLU2_OP410_030 := [[-129.18,-85.76,185.33],[0.128544,-0.701387,0.295212,-0.635911],[-1,1,1,0],[9E+09,9E+09,9E+09,9E+09,9E+09,9E+09]];
    PERS robtarget pLU2_OP410_040 := [[-125.52,-69.68,192.94],[0.128541,-0.701386,0.295209,-0.635914],[-1,1,1,0],[9E+09,9E+09,9E+09,9E+09,9E+09,9E+09]];
    PERS robtarget pLU2_OP410_050 := [[-137.77,-69.68,192.93],[0.128541,-0.701388,0.295211,-0.635911],[-1,1,1,0],[9E+09,9E+09,9E+09,9E+09,9E+09,9E+09]];
    PERS robtarget pLU2_OP410_060 := [[-127.69,-20.57,203.99],[0.0880921,-0.731082,0.0960536,-0.669726],[-1,1,0,0],[9E+09,9E+09,9E+09,9E+09,9E+09,9E+09]];
    PERS robtarget pLU2_OP410_070 := [[-117.15,-20.58,203.97],[0.0880955,-0.731083,0.0960578,-0.669723],[-1,1,0,0],[9E+09,9E+09,9E+09,9E+09,9E+09,9E+09]];
    PERS robtarget pLU2_OP410_080 := [[-110.59,-23.45,168.72],[0.0880952,-0.731084,0.0960575,-0.669723],[-1,1,0,0],[9E+09,9E+09,9E+09,9E+09,9E+09,9E+09]];
    PERS robtarget pLU2_OP410_090 := [[-109.13,-23.45,163.37],[0.0881014,-0.731094,0.0960692,-0.669709],[-1,1,0,0],[9E+09,9E+09,9E+09,9E+09,9E+09,9E+09]];
    PERS robtarget pLU2_OP410_100 := [[-103.49,-23.45,150.78],[0.0880987,-0.731093,0.0960653,-0.669711],[-1,1,0,0],[9E+09,9E+09,9E+09,9E+09,9E+09,9E+09]];
    PERS robtarget pLU2_OP410_110 := [[-45.32,-19.48,48.40],[0.0880965,-0.731091,0.0960606,-0.669714],[-1,1,0,0],[9E+09,9E+09,9E+09,9E+09,9E+09,9E+09]];
    PERS robtarget pLU2_OP410_120 := [[-55.15,-19.48,37.59],[0.0881002,-0.731095,0.0960664,-0.669709],[-1,1,0,0],[9E+09,9E+09,9E+09,9E+09,9E+09,9E+09]];
    PERS robtarget pLU2_OP410_130 := [[-257.91,-19.48,-4.69],[0.0881005,-0.731094,0.096068,-0.669709],[-1,1,0,0],[9E+09,9E+09,9E+09,9E+09,9E+09,9E+09]];
    !New
    PERS robtarget pL0:=[[0,0,0],[0,0,0,0],[0,0,0,0],[9E+09,9E+09,9E+09,9E+09,9E+09,9E+09]];







PROC A1_Change()
    R_Home;
    !Approach to the position
 MoveJ pLAppChange10_,vWithPart,z50,tGripp_1;
 MoveJ pLAppChange9_,vWithPart,z50,tGripp_1;
 MoveJ pLAppChange8_,vWithPart,z50,tGripp_1;
 MoveJ pLAppChange7_,vWithPart,z50,tGripp_1;
 MoveJ pLAppChange6_,vWithPart,z50,tGripp_1;
 MoveJ pLAppChange5_,vWithPart,z50,tGripp_1;
 MoveJ pLAppChange4_,vWithPart,z50,tGripp_1;
 MoveJ pLAppChange3_,vWithPart,z50,tGripp_1;
 MoveJ pLAppChange2_,vWithPart,z50,tGripp_1;
 MoveJ pLAppChange1_,vWithPart,z50,tGripp_1;
    R_Home;
    !
ENDPROC


ENDMODULE
